// TwinCAT 3 PLC project lamppuprosessi
// ProgramVersion: 3.1.4026.27
// libraries:
//   Tc2_Standard, * (Beckhoff Automation GmbH)
//   Tc2_System, * (Beckhoff Automation GmbH)
//   Tc3_IotBase, * (Beckhoff Automation GmbH)
//   Tc3_Module, * (Beckhoff Automation GmbH)
// project tree:
//   GVLs/ GVL.TcGVL
//   / PlcTask.TcTTO
//   POUs/ MAIN.TcPOU, MQTTpublisher.TcPOU, MQTTsubscriber.TcPOU, PIcontroller.TcPOU
// real-time tasks:
//   TASK PlcTask: cycle T#10ms, priority 20, ADS port 350
// I/O:
//   DEVICE Device 1 (EtherCAT), AmsNetId 5.159.149.51.2.1
//     Term 1 (EK1200) [EK1200-7000 EtherCAT Power supply (1,5A E-Bus)]
//       Term 2 (EL3202) [EL3202 2Ch. Ana. Input PT100 (RTD)]
//       Term 3 (EL4102) [EL4102 2Ch. Ana. Output  0-10V, 16bit]
//       Term 4 (EL9011) [EL9011 End Terminal]
//   DEVICE Device 2 (NOV-DP-RAM)
//   DEVICE Device 3 (CX7000), AmsNetId 5.159.149.51.4.1
//     Term 1 (CX7028) [CX7028-0000-0118]
//       modules: Module 1 (DIO_2x), Module 3 (DIO_2x), Module 5 (DI_2x), Module 7 (DI_2x)
// variable links:
//   lamppuprosessi/lamppuprosessi Instance <-> Device 1 (EtherCAT)/Term 1 (EK1200)/Term 2 (EL3202)
//     PlcTask Inputs/GVL.iPT100rawdata <-> RTD Inputs Channel 1/Value
//   lamppuprosessi/lamppuprosessi Instance <-> Device 1 (EtherCAT)/Term 1 (EK1200)/Term 3 (EL4102)
//     PlcTask Outputs/GVL.iLampPower <-> Channel 1/Output

CONFIGURATION lamppuprosessi
    RESOURCE PLC ON TwinCAT3
        TASK PlcTask(INTERVAL := T#10ms, PRIORITY := 20);
        PROGRAM MAIN WITH PlcTask : MAIN;
    END_RESOURCE
END_CONFIGURATION

// ---- GVLs/GVL.TcGVL
{attribute 'qualified_only'}
VAR_GLOBAL
	iPT100rawdata AT %I* : INT;
	iLampPower	AT %Q* : INT;
END_VAR

// ---- POUs/MAIN.TcPOU
PROGRAM MAIN
VAR
	Controller      : PIcontroller;
	Lamp_temp		: REAL;				// Lamp temperature in Celsius
	Temp_setpoint	: REAL := 30;		// write values to change the setpoint
	
	PI_Kp			: REAL;				// Gain 
	PI_Ki			: REAL;				// Integral
	
	fbMQTTPublisher : MQTTpublisher;
	fbSubscriber	:MQTTsubscriber;
END_VAR

// PI Controller
Controller(		MeasuredValue := GVL.iPT100rawdata,
				Setpoint 	  := Temp_setpoint,
				Kp			  := PI_Kp,
				Ki			  := PI_Ki,);

				
// Scales the data from the PT100 Sensor to Celsius.	
Lamp_temp := INT_TO_REAL(GVL.iPT100rawdata) / 10.0;

// Scales the PI controller 0-100 value to an analog 16 bit value 0-32767.
GVL.iLampPower := REAL_TO_INT(Controller.ControlValue * 327.67);

// Publishes the lamp temperature to MQTT once per second
fbMQTTPublisher(fValue := Lamp_temp);

// Receives setpoint, Kp and Ki over MQTT
fbSubscriber(fSetpoint := Temp_setpoint, fKp := PI_Kp, fKi := PI_Ki);

END_PROGRAM

// ---- POUs/PIcontroller.TcPOU
FUNCTION_BLOCK PIcontroller

VAR_INPUT
	MeasuredValue			: REAL;
	SetPoint				: REAL;
    Kp 						: REAL;          
    Ki 						: REAL;	
END_VAR

VAR_OUTPUT
	ControlValue			: REAL;
END_VAR

VAR
	ProcessVariable 		: REAL;  			(* Current process value *)
    TimeCycle 				: REAL:=0.01;       (* Cycle time in seconds *)
    ControlOutput 			: REAL;          	(* PID controller output *)
    Error 					: REAL;            	(* Difference between SetPoint and ProcessVariable *)
    Integral 				: REAL;         	(* Integral accumulator *)
    Derivative 				: REAL;       		(* Derivative term *)
    PrevError 				: REAL;        		(* Error from the previous cycle *)
	PrevSetPoint 			: REAL := 0.0;
END_VAR

// PI CONTROLLER

ProcessVariable:=MeasuredValue;
 
IF SetPoint <> PrevSetPoint THEN // Integral value resets to zero everytime the setpoint is changed to avoid integral windup.
    Integral := 0.0;
    PrevSetPoint := SetPoint;
END_IF

Error := (SetPoint * 10) - ProcessVariable; // Error = How far away from the setpoint the temperature is.
	
    IF (ControlOutput = ControlValue) OR 		// Integral value won't change unless these conditions are met. This is to avoid windup.
       (ControlOutput > 100.0 AND Error < 0.0) OR 
       (ControlOutput < 0.0 AND Error > 0.0) THEN
	   
	   Integral := Integral + (Ki * Error * TimeCycle);
	END_IF
    
ControlOutput := (Kp * Error) + (Ki * Integral); // PI controller math
	
ControlValue := LIMIT(0,ControlOutput,100);	// Limits the control to only go from 0 to 100

END_FUNCTION_BLOCK

// ---- POUs/MQTTpublisher.TcPOU
FUNCTION_BLOCK MQTTpublisher
VAR_INPUT
	bEnable     : BOOL := TRUE;
    sHostName   : STRING(255) := '192.168.0.100';   // The PC's IP on the PLC network
    nHostPort   : UINT := 1883;
    sClientId   : STRING(255) := 'CX7000-publisher';
    sTopic      : STRING(255) := 'plc/pid/temp';
    fValue      : REAL;                              // Value to publish
    tInterval   : TIME := T#1S;                      // Publish interval
END_VAR

VAR_OUTPUT
	 bConnected  : BOOL;
    bError      : BOOL;
    hrErrorCode : HRESULT;
END_VAR

VAR
	fbMqttClient : FB_IotMqttClient;
    fbTimer      : TON;
    bInit        : BOOL := TRUE;
    sPayload     : STRING(255);
END_VAR

// Set the connection parameters once
IF bInit THEN
    bInit := FALSE;
    fbMqttClient.sHostName := sHostName;
    fbMqttClient.nHostPort := nHostPort;
    fbMqttClient.sClientId := sClientId;
END_IF

// Must be called every cycle: keeps the connection alive
fbMqttClient.Execute(bEnable);

bConnected  := fbMqttClient.bConnected;
bError      := fbMqttClient.bError;
hrErrorCode := fbMqttClient.hrErrorCode;

// Publish once per interval while connected
fbTimer(IN := bConnected AND NOT fbTimer.Q, PT := tInterval);

IF fbTimer.Q THEN
    sPayload := REAL_TO_STRING(fValue);
    fbMqttClient.Publish(
        sTopic       := sTopic,
        pPayload     := ADR(sPayload),
        nPayloadSize := INT_TO_UDINT(LEN(sPayload)),
        eQoS         := TcIotMqttQos.AtMostOnceDelivery,
        bRetain      := FALSE,
        bQueue       := FALSE);
END_IF

END_FUNCTION_BLOCK

// ---- POUs/MQTTsubscriber.TcPOU
FUNCTION_BLOCK MQTTsubscriber
VAR_INPUT
    bEnable     : BOOL := TRUE;
    sHostName   : STRING(255) := '192.168.0.100';   // The PC's IP on the PLC network
    nHostPort   : UINT := 1883;
    sClientId   : STRING(255) := 'CX7000-subscriber';      // Must differ from the publisher's
    sTopicSub   : STRING(255) := 'plc/pid/#';
END_VAR
VAR_OUTPUT
    bConnected  : BOOL;
    bSubscribed : BOOL;
    bError      : BOOL;
    hrErrorCode : HRESULT;
    nRxCount    : UDINT;                             // Number of messages received (for debugging)
END_VAR
VAR_IN_OUT
    fSetpoint   : REAL;                              // Only changed when a message arrives
    fKp         : REAL;
    fKi         : REAL;
END_VAR
VAR
    fbMqttClient   : FB_IotMqttClient;
    fbMessageQueue : FB_IotMqttMessageQueue;
    fbMessage      : FB_IotMqttMessage;
    bInit          : BOOL := TRUE;
    sTopicRcv      : STRING(255);
    sPayloadRcv    : STRING(255);
END_VAR

// Set the connection parameters once
IF bInit THEN
    bInit := FALSE;
    fbMqttClient.sHostName      := sHostName;
    fbMqttClient.nHostPort      := nHostPort;
    fbMqttClient.sClientId      := sClientId;
    fbMqttClient.ipMessageQueue := fbMessageQueue;
END_IF

// Must be called every cycle
fbMqttClient.Execute(bEnable);

bConnected  := fbMqttClient.bConnected;
bError      := fbMqttClient.bError;
hrErrorCode := fbMqttClient.hrErrorCode;

IF bConnected THEN
    // Subscribe once after connecting
    IF NOT bSubscribed THEN
        bSubscribed := fbMqttClient.Subscribe(sTopic := sTopicSub,
                                              eQoS   := TcIotMqttQos.AtMostOnceDelivery);
    END_IF

    // Handle all received messages
    WHILE fbMessageQueue.nQueuedMessages > 0 DO
        IF fbMessageQueue.Dequeue(fbMessage := fbMessage) THEN
            fbMessage.GetTopic(pTopic := ADR(sTopicRcv), nTopicSize := SIZEOF(sTopicRcv));
            fbMessage.GetPayload(pPayload            := ADR(sPayloadRcv),
                                 nPayloadSize        := SIZEOF(sPayloadRcv),
                                 bSetNullTermination := TRUE);
            nRxCount := nRxCount + 1;

            IF sTopicRcv = 'plc/pid/setpoint' THEN
                fSetpoint := STRING_TO_REAL(sPayloadRcv);
            ELSIF sTopicRcv = 'plc/pid/kp' THEN
                fKp := STRING_TO_REAL(sPayloadRcv);
            ELSIF sTopicRcv = 'plc/pid/ki' THEN
                fKi := STRING_TO_REAL(sPayloadRcv);
            END_IF
            // plc/pid/temp (the PLC's own publication) is ignored
        END_IF
    END_WHILE
ELSE
    bSubscribed := FALSE;   // Subscribe again after reconnecting
END_IF

END_FUNCTION_BLOCK
